// TIA Portal V19 export
DATA_BLOCK "AI_INST_RANG"   // DB80
{ S7_Optimized_Access := 'FALSE' }
   VAR RETAIN
      R1_TT01 : Struct
         MIN : Real := -50.0;
         MAX : Real := 200.0;
      END_STRUCT;
      R1_TT02 : Struct
         MIN : Real := -50.0;
         MAX : Real := 200.0;
      END_STRUCT;
      R1_TT03 : Struct
         MIN : Real := -50.0;
         MAX : Real := 200.0;
      END_STRUCT;
      R2_TT01 : Struct
         MIN : Real := -50.0;
         MAX : Real := 200.0;
      END_STRUCT;
      R2_TT02 : Struct
         MIN : Real := -50.0;
         MAX : Real := 200.0;
      END_STRUCT;
      R2_TT03 : Struct
         MIN : Real := -50.0;
         MAX : Real := 200.0;
      END_STRUCT;
      R3_TT01 : Struct
         MIN : Real := -50.0;
         MAX : Real := 200.0;
      END_STRUCT;
      R3_TT02 : Struct
         MIN : Real := -50.0;
         MAX : Real := 200.0;
      END_STRUCT;
      R3_TT03 : Struct
         MIN : Real := -50.0;
         MAX : Real := 200.0;
      END_STRUCT;
      R4_TT01 : Struct
         MIN : Real := -50.0;
         MAX : Real := 200.0;
      END_STRUCT;
      R4_TT02 : Struct
         MIN : Real := -50.0;
         MAX : Real := 200.0;
      END_STRUCT;
      R4_TT03 : Struct
         MIN : Real := -50.0;
         MAX : Real := 200.0;
      END_STRUCT;
      R5_TT01 : Struct
         MIN : Real := -50.0;
         MAX : Real := 200.0;
      END_STRUCT;
      R5_TT02 : Struct
         MIN : Real := -50.0;
         MAX : Real := 200.0;
      END_STRUCT;
      R5_TT03 : Struct
         MIN : Real := -50.0;
         MAX : Real := 200.0;
      END_STRUCT;
      R6_TT01 : Struct
         MIN : Real := -50.0;
         MAX : Real := 200.0;
      END_STRUCT;
      R6_TT02 : Struct
         MIN : Real := -50.0;
         MAX : Real := 200.0;
      END_STRUCT;
      R6_TT03 : Struct
         MIN : Real := -50.0;
         MAX : Real := 200.0;
      END_STRUCT;
      R7_TT01 : Struct
         MIN : Real := -50.0;
         MAX : Real := 200.0;
      END_STRUCT;
      R7_TT02 : Struct
         MIN : Real := -50.0;
         MAX : Real := 200.0;
      END_STRUCT;
      R7_TT03 : Struct
         MIN : Real := -50.0;
         MAX : Real := 200.0;
      END_STRUCT;
      R8_TT01 : Struct
         MIN : Real := -50.0;
         MAX : Real := 200.0;
      END_STRUCT;
      R8_TT02 : Struct
         MIN : Real := -50.0;
         MAX : Real := 200.0;
      END_STRUCT;
      R8_TT03 : Struct
         MIN : Real := -50.0;
         MAX : Real := 200.0;
      END_STRUCT;
      R9_TT01 : Struct
         MIN : Real := -50.0;
         MAX : Real := 200.0;
      END_STRUCT;
      R9_TT02 : Struct
         MIN : Real := -50.0;
         MAX : Real := 200.0;
      END_STRUCT;
      R9_TT03 : Struct
         MIN : Real := -50.0;
         MAX : Real := 200.0;
      END_STRUCT;
      R10_TT01 : Struct
         MIN : Real := -50.0;
         MAX : Real := 200.0;
      END_STRUCT;
      R10_TT02 : Struct
         MIN : Real := -50.0;
         MAX : Real := 200.0;
      END_STRUCT;
      R10_TT03 : Struct
         MIN : Real := -50.0;
         MAX : Real := 200.0;
      END_STRUCT;
      R11_TT01 : Struct
         MIN : Real := -50.0;
         MAX : Real := 200.0;
      END_STRUCT;
      R11_TT02 : Struct
         MIN : Real := -50.0;
         MAX : Real := 200.0;
      END_STRUCT;
      R11_TT03 : Struct
         MIN : Real := -50.0;
         MAX : Real := 200.0;
      END_STRUCT;
      R12_TT01 : Struct
         MIN : Real := -50.0;
         MAX : Real := 200.0;
      END_STRUCT;
      R12_TT02 : Struct
         MIN : Real := -50.0;
         MAX : Real := 200.0;
      END_STRUCT;
      R12_TT03 : Struct
         MIN : Real := -50.0;
         MAX : Real := 200.0;
      END_STRUCT;
      R13_TT01 : Struct
         MIN : Real := -50.0;
         MAX : Real := 200.0;
      END_STRUCT;
      R13_TT02 : Struct
         MIN : Real := -50.0;
         MAX : Real := 200.0;
      END_STRUCT;
      R13_TT03 : Struct
         MIN : Real := -50.0;
         MAX : Real := 200.0;
      END_STRUCT;
      R14_TT01 : Struct
         MIN : Real := -50.0;
         MAX : Real := 200.0;
      END_STRUCT;
      R14_TT02 : Struct
         MIN : Real := -50.0;
         MAX : Real := 200.0;
      END_STRUCT;
      R14_TT03 : Struct
         MIN : Real := -50.0;
         MAX : Real := 200.0;
      END_STRUCT;
      R15_TT01 : Struct
         MIN : Real := -50.0;
         MAX : Real := 200.0;
      END_STRUCT;
      R15_TT02 : Struct
         MIN : Real := -50.0;
         MAX : Real := 200.0;
      END_STRUCT;
      R15_TT03 : Struct
         MIN : Real := -50.0;
         MAX : Real := 200.0;
      END_STRUCT;
      R16_TT01 : Struct
         MIN : Real := -50.0;
         MAX : Real := 200.0;
      END_STRUCT;
      R16_TT02 : Struct
         MIN : Real := -50.0;
         MAX : Real := 200.0;
      END_STRUCT;
      R16_TT03 : Struct
         MIN : Real := -50.0;
         MAX : Real := 200.0;
      END_STRUCT;
      R17_TT01 : Struct
         MIN : Real := -50.0;
         MAX : Real := 200.0;
      END_STRUCT;
      R17_TT02 : Struct
         MIN : Real := -50.0;
         MAX : Real := 200.0;
      END_STRUCT;
      R17_TT03 : Struct
         MIN : Real := -50.0;
         MAX : Real := 200.0;
      END_STRUCT;
      R18_TT01 : Struct
         MIN : Real := -50.0;
         MAX : Real := 200.0;
      END_STRUCT;
      R18_TT02 : Struct
         MIN : Real := -50.0;
         MAX : Real := 200.0;
      END_STRUCT;
      R18_TT03 : Struct
         MIN : Real := -50.0;
         MAX : Real := 200.0;
      END_STRUCT;
      CHS_TT01 : Struct
         MIN : Real := -50.0;
         MAX : Real := 200.0;
      END_STRUCT;
      CHS_TT02 : Struct
         MIN : Real := -50.0;
         MAX : Real := 200.0;
      END_STRUCT;
      CHS_TT03 : Struct
         MIN : Real := -50.0;
         MAX : Real := 200.0;
      END_STRUCT;
      CHS_TT04 : Struct
         MIN : Real := -50.0;
         MAX : Real := 200.0;
      END_STRUCT;
      CHS_MGLT : Struct
         MIN : Real := -50.0;
         MAX : Real := 200.0;
      END_STRUCT;
      CH_PT01 : Struct
         MIN : Real := -50.0;
         MAX : Real := 200.0;
      END_STRUCT;
      SMHS_TT01 : Struct
         MIN : Real := -50.0;
         MAX : Real := 200.0;
      END_STRUCT;
      SMCS_TT02 : Struct
         MIN : Real := -50.0;
         MAX : Real := 200.0;
      END_STRUCT;
      SMCHS_TT03 : Struct
         MIN : Real := -50.0;
         MAX : Real := 200.0;
      END_STRUCT;
      SMUCHS_TT04 : Struct
         MIN : Real := -50.0;
         MAX : Real := 200.0;
      END_STRUCT;
      NMHS_TT01 : Struct
         MIN : Real := -50.0;
         MAX : Real := 200.0;
      END_STRUCT;
      NMCS_TT02 : Struct
         MIN : Real := -50.0;
         MAX : Real := 200.0;
      END_STRUCT;
      NMCHS_TT03 : Struct
         MIN : Real := -50.0;
         MAX : Real := 200.0;
      END_STRUCT;
      NMUCHS_TT04 : Struct
         MIN : Real := -50.0;
         MAX : Real := 200.0;
      END_STRUCT;
      SMHS_PT01 : Struct
         MIN : Real := -50.0;
         MAX : Real := 200.0;
      END_STRUCT;
      SMCS_PT02 : Struct
         MIN : Real := -50.0;
         MAX : Real := 200.0;
      END_STRUCT;
      SMCHS_PT03 : Struct
         MIN : Real := -50.0;
         MAX : Real := 200.0;
      END_STRUCT;
      SMUCHS_PT04 : Struct
         MIN : Real := -50.0;
         MAX : Real := 200.0;
      END_STRUCT;
      NMHS_PT01 : Struct
         MIN : Real := -50.0;
         MAX : Real := 200.0;
      END_STRUCT;
      NMCS_PT02 : Struct
         MIN : Real := -50.0;
         MAX : Real := 200.0;
      END_STRUCT;
      NMCHS_PT03 : Struct
         MIN : Real := -50.0;
         MAX : Real := 200.0;
      END_STRUCT;
      NMUCHS_PT04 : Struct
         MIN : Real := -50.0;
         MAX : Real := 200.0;
      END_STRUCT;
      CS_TT01 : Struct
         MIN : Real := -50.0;
         MAX : Real := 200.0;
      END_STRUCT;
      CS_TT02 : Struct
         MIN : Real := -50.0;
         MAX : Real := 200.0;
      END_STRUCT;
      CS_TT03 : Struct
         MIN : Real := -50.0;
         MAX : Real := 200.0;
      END_STRUCT;
      CS_TT04 : Struct
         MIN : Real := -50.0;
         MAX : Real := 200.0;
      END_STRUCT;
      CS_MGLT : Struct
         MIN : Real := -50.0;
         MAX : Real := 200.0;
      END_STRUCT;
      UCHS_TT01 : Struct
         MIN : Real := -50.0;
         MAX : Real := 200.0;
      END_STRUCT;
      UCHS_TT02 : Struct
         MIN : Real := -50.0;
         MAX : Real := 200.0;
      END_STRUCT;
      UCHS_TT03 : Struct
         MIN : Real := -50.0;
         MAX : Real := 200.0;
      END_STRUCT;
      UCHS_TT04 : Struct
         MIN : Real := -50.0;
         MAX : Real := 200.0;
      END_STRUCT;
      UCHS_MGLT : Struct
         MIN : Real := -50.0;
         MAX : Real := 200.0;
      END_STRUCT;
      HS_TT01 : Struct
         MIN : Real := -50.0;
         MAX : Real := 200.0;
      END_STRUCT;
      HS_TT02 : Struct
         MIN : Real := -50.0;
         MAX : Real := 200.0;
      END_STRUCT;
      HS_TT03 : Struct
         MIN : Real := -50.0;
         MAX : Real := 200.0;
      END_STRUCT;
      HS_MGLT : Struct
         MIN : Real := -50.0;
         MAX : Real := 200.0;
      END_STRUCT;
      "AI_A/SCRB_001_PH01" : Struct
         MIN : Real := -50.0;
         MAX : Real := 200.0;
      END_STRUCT;
      "AI_A/SCRB_002_PH01" : Struct
         MIN : Real := -50.0;
         MAX : Real := 200.0;
      END_STRUCT;
      "A/VP_01_APT01" : Struct
         MIN : Real := -50.0;
         MAX : Real := 200.0;
      END_STRUCT;
      "A/VP_02_APT01" : Struct
         MIN : Real := -50.0;
         MAX : Real := 200.0;
      END_STRUCT;
      "A/ANFD_001_APT01" : Struct
         MIN : Real := -50.0;
         MAX : Real := 200.0;
      END_STRUCT;
      "A/ANFD_002_APT01" : Struct
         MIN : Real := -50.0;
         MAX : Real := 200.0;
      END_STRUCT;
      "A/ANFD_003_APT01" : Struct
         MIN : Real := -50.0;
         MAX : Real := 200.0;
      END_STRUCT;
      "A/ANFD_004_APT01" : Struct
         MIN : Real := -50.0;
         MAX : Real := 200.0;
      END_STRUCT;
      "A/ANFD_001_TT01" : Struct
         MIN : Real := -50.0;
         MAX : Real := 200.0;
      END_STRUCT;
      "A/ANFD_002_TT01" : Struct
         MIN : Real := -50.0;
         MAX : Real := 200.0;
      END_STRUCT;
      "A/ANFD_003_TT01" : Struct
         MIN : Real := -50.0;
         MAX : Real := 200.0;
      END_STRUCT;
      "A/ANFD_004_TT01" : Struct
         MIN : Real := -50.0;
         MAX : Real := 200.0;
      END_STRUCT;
      RCVD_001_APT01 : Struct
         MIN : Real := -50.0;
         MAX : Real := 200.0;
      END_STRUCT;
      RCVD_002_APT01 : Struct
         MIN : Real := -50.0;
         MAX : Real := 200.0;
      END_STRUCT;
      RCVD_001_TT01 : Struct
         MIN : Real := -50.0;
         MAX : Real := 200.0;
      END_STRUCT;
      RCVD_002_TT01 : Struct
         MIN : Real := -50.0;
         MAX : Real := 200.0;
      END_STRUCT;
      "AI_A/VTD_001_APT01" : Struct
         MIN : Real := -50.0;
         MAX : Real := 200.0;
      END_STRUCT;
      "AI_A/VTD_002_APT01" : Struct
         MIN : Real := -50.0;
         MAX : Real := 200.0;
      END_STRUCT;
      "AI_A/VTD_001_TT01" : Struct
         MIN : Real := -50.0;
         MAX : Real := 200.0;
      END_STRUCT;
      "AI_A/VTD_002_TT01" : Struct
         MIN : Real := -50.0;
         MAX : Real := 200.0;
      END_STRUCT;
      "AI_A/TD_001_TT01" : Struct
         MIN : Real := -50.0;
         MAX : Real := 200.0;
      END_STRUCT;
      "AI_A/TD_002_TT01" : Struct
         MIN : Real := -50.0;
         MAX : Real := 200.0;
      END_STRUCT;
   END_VAR
BEGIN
END_DATA_BLOCK
